TYPE ST_CamParam :
STRUCT
	bCamLoad: BOOL;
	bPeriodic: BOOL;
	nElements: UINT;
	nBuffNum: UINT;
	nPointType: UINT;
	aCamBuffer: ARRAY[0..9] OF ST_CamXYVA;
END_STRUCT
END_TYPE

(* stored: Version 1.1.0.1, ProductVersion 3.1.4024.12
   DUT ST_CamParam: Id {8dff8ca0-22b0-4cf5-9ebe-b6027cba8191} *)
